FUNCTION_BLOCK R1 (* Basic Function Block Type *)
  (* Standard: 61499-2 *)
  (* Version 0.0, 10/11/2026, lizar, nxtControl GmBH, Template *)
  PACKAGE Main;
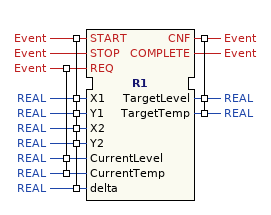
  EVENT_INPUT
    START WITH X1, Y1, X2, Y2, delta; (* Normal Execution Request *)
    STOP;
    REQ WITH CurrentLevel, CurrentTemp;
  END_EVENT
  EVENT_OUTPUT
    CNF WITH TargetLevel, TargetTemp; (* Execution Confirmation *)
    COMPLETE;
  END_EVENT
  VAR_INPUT
    X1 : REAL; (* Input event qualifier *)
    Y1 : REAL;
    X2 : REAL;
    Y2 : REAL;
    CurrentLevel : REAL;
    CurrentTemp : REAL;
    delta : REAL;
  END_VAR
  VAR_OUTPUT
    TargetLevel : REAL;
    TargetTemp : REAL;
  END_VAR
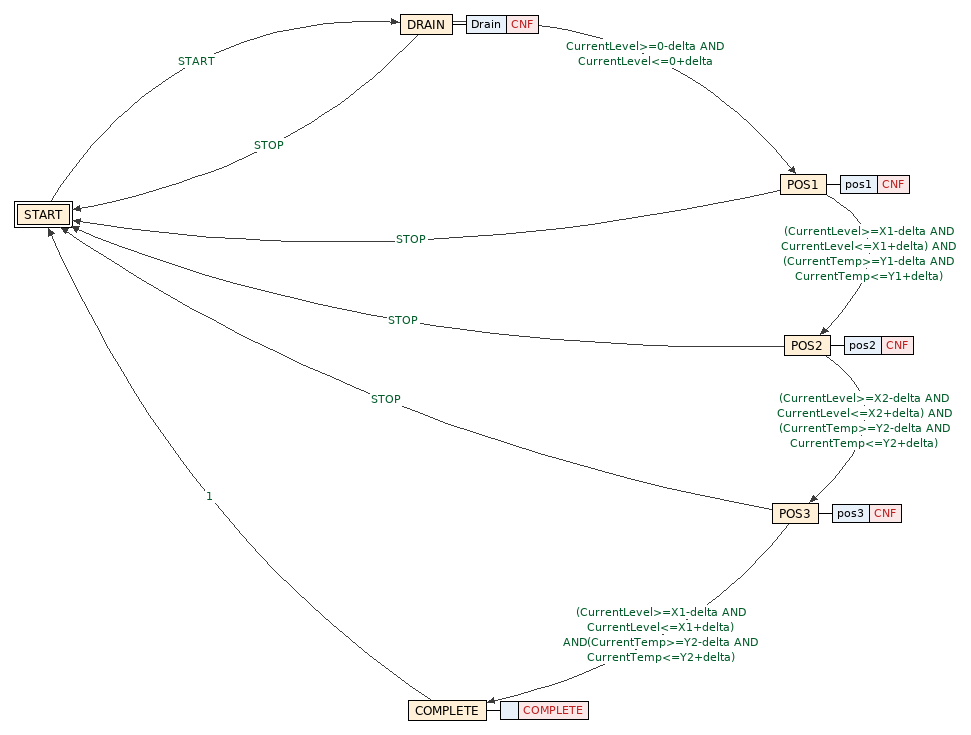
  EC_STATES
    START; (* Initial State *)
    DRAIN : Drain -> CNF;
    POS1 : pos1 -> CNF;
    POS2 : pos2 -> CNF;
    POS3 : pos3 -> CNF;
    COMPLETE : -> COMPLETE;
  END_STATES
  EC_TRANSITIONS
    START TO DRAIN := START;
    DRAIN TO POS1 := CurrentLevel>=0-delta AND CurrentLevel<=0+delta;
    POS1 TO POS2 := (CurrentLevel>=X1-delta AND CurrentLevel<=X1+delta) AND (CurrentTemp>=Y1-delta AND CurrentTemp<=Y1+delta);
    POS2 TO POS3 := (CurrentLevel>=X2-delta AND CurrentLevel<=X2+delta) AND (CurrentTemp>=Y2-delta AND CurrentTemp<=Y2+delta);
    POS3 TO COMPLETE := (CurrentLevel>=X1-delta AND CurrentLevel<=X1+delta) AND(CurrentTemp>=Y2-delta AND CurrentTemp<=Y2+delta);
    COMPLETE TO START := 1;
    DRAIN TO START := STOP;
    POS1 TO START := STOP;
    POS2 TO START := STOP;
    POS3 TO START := STOP;
  END_TRANSITIONS
  ALGORITHM Drain IN ST:
TargetLevel:= 0;
TargetTemp := 0;
  END_ALGORITHM
  ALGORITHM pos1 IN ST:
TargetLevel:= X1;
TargetTemp := Y1;
  END_ALGORITHM
  ALGORITHM pos2 IN ST:
TargetLevel:= X2;
TargetTemp := Y2;
  END_ALGORITHM
  ALGORITHM pos3 IN ST:
TargetLevel:= X1;
  END_ALGORITHM
END_FUNCTION_BLOCK
